Yaskawa INFORM job: SQUARE.JBI

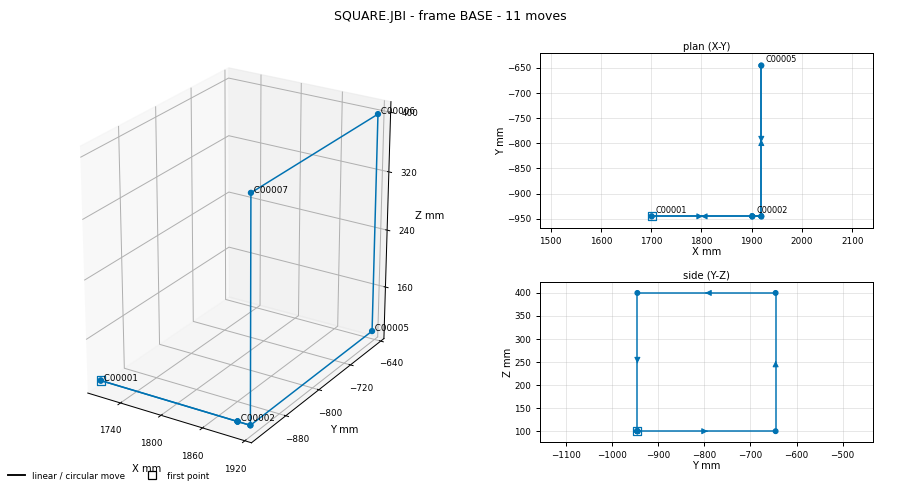
[picture p0: tool path of SQUARE.JBI in frame BASE, 11 of 12 moves have a stored position in this frame; points joined in program order, loops and branches not executed]
/JOB
//NAME SQUARE
//POS
///NPOS 12,0,0,0,0,0
///TOOL 9
///POSTYPE PULSE
///PULSE
C00000=-35,27,-31,39,65,-109
///TOOL 9
///POSTYPE BASE
///RECTAN
///RCONF 1,0,0,0,0,0,0,0
C00001=1701.000,-945.302,100.000,-90.00,-0.00,-90.00
C00002=1901.000,-945.302,100.000,-90.00,-0.00,-90.00
C00003=1901.000,-945.302,100.000,-90.00,-0.00,-90.00
C00004=1919.000,-945.302,100.000,-90.00,-0.00,-90.00
C00005=1919.000,-645.302,100.000,-90.00,-0.00,-90.00
C00006=1919.000,-645.302,400.000,-90.00,-0.00,-90.00
C00007=1919.000,-945.302,400.000,-90.00,-0.00,-90.00
C00008=1919.000,-945.302,100.000,-90.00,-0.00,-90.00
C00009=1901.000,-945.302,100.000,-90.00,-0.00,-90.00
C00010=1901.000,-945.302,100.000,-90.00,-0.00,-90.00
C00011=1701.000,-945.302,100.000,-90.00,-0.00,-90.00
//INST
///DATE 2026/10/26 01:19
///COMM Generated using RoboDK
///ATTR SC,RW,RJ
///GROUP1 RB1
NOP
'Using Tool1 (targets wrt base
'):
'1921.0,-795.3,250.0,90.0,0.0,
'-90.0
'Setting Tool 9 (BALL END - 10
'MM):
SETE P00095 (1) 0
SETE P00095 (2) 0
SETE P00095 (3) 85000
SETE P00095 (4) 0
SETE P00095 (5) 0
SETE P00095 (6) 0
SETTOOL TL#(9) P00095
'hide USER - ENGRAVE - 30 DEG
'POINT END
'show BALL END - 10MM
MSG "/ ALPHACAM DRAWING FILE -"
MSG " ROBOTAPT"
MSG "/ NC CODE FILE - ROBOTAPT"
MSG ".apt"
MSG "/ POST-PROCESSED FOR APT-"
MSG "CL DATA"
MSG "/ CREATED - 26 NOV 18"
MSG "/ PROGRAMMED BY ALPHACAM"
MSG "/ BALL END - 10MM"
MOVJ C00000 VJ=50.00
MOVL C00001 V=1000.0
MOVL C00002 V=1000.0
CALL JOB:SPINDLE
MOVL C00003 V=1000.0
MOVL C00004 V=160.0
MOVL C00005 V=160.0
MOVL C00006 V=160.0
MOVL C00007 V=160.0
MOVL C00008 V=160.0
MOVL C00009 V=1000.0
CALL JOB:SPINDLE
MOVL C00010 V=1000.0
MOVL C00011 V=1000.0
END
